// TIA Portal V21 export
// export: Created 2026-08-21T20:18:53.1493152Z, ExportSetting None, DisplayName Totally Integrated Automation Portal, DisplayVersion V21, DisplayName STEP 7 Professional, DisplayVersion V21, DisplayName STEP 7 Safety, DisplayVersion V21, DisplayName Tech WebApplication, DisplayVersion V21, DisplayName WinCC Basic/Comfort/Advanced, DisplayVersion V21, DisplayName WinCC Professional, DisplayVersion V21, DisplayName WinCC Unified, DisplayVersion V21
FUNCTION_BLOCK "ConfigurationParameters"   // FB1710, SCL
TITLE = ConfigurationParameters
{ S7_Optimized_Access := 'TRUE' }
AUTHOR : Siemens AG
FAMILY : ServiceControl
VERSION : 1.0
// Providing of the MTP-Interface and the number of parameters of each configuration parameter type
// stored: MemoryReserve 100, SetENOAutomatically false
   VAR
      MTPAnalog { S7_SetPoint := 'True'} : Array[0..#NUMBER_PARAMETERS_ANALOG] of "UDT_MTP_AnaServParam";
      MTPDigital { S7_SetPoint := 'True'} : Array[0..#NUMBER_PARAMETERS_DIGITAL] of "UDT_MTP_DIntServParam";
      MTPBinary { S7_SetPoint := 'True'} : Array[0..#NUMBER_PARAMETERS_BINARY] of "UDT_MTP_BinServParam";
      MTPString { S7_SetPoint := 'True'} : Array[0..#NUMBER_PARAMETERS_STRING] of "UDT_MTP_StringServParam";
   END_VAR
   VAR CONSTANT
      NUMBER_PARAMETERS_ANALOG : Int := 0;
      NUMBER_PARAMETERS_DIGITAL : Int := 0;
      NUMBER_PARAMETERS_BINARY : Int := 1;
      NUMBER_PARAMETERS_STRING : Int := 0;
   END_VAR
BEGIN
   REGION Block Info Header
     //===============================================================================
     // Siemens AG / (c)Copyright 2021
     //-------------------------------------------------------------------------------
     // Title:            ConfigurationParameters
     // Comment/Function: Providing of the MTP-Interface and the number of parameters of each configuration parameter type
     // Library/Family:   ServiceControl
     // Author:           Siemens AG
     // Tested with:      S7-PLCSIM Advanced 4.0
     // Engineering:      TIA Portal V17
     // Restrictions:     MTP
     // Requirements:     PLC (S7-1200 / S7-1500)
     //-------------------------------------------------------------------------------
     // Change log table:
     // Version  | Date       | Expert in charge        | Changes applied
     //----------|------------|-------------------------|-----------------------------
     // 01.00.00 | 02.09.2021 | Michael Schlosser       | First released version
     // 01.00.01 | 07.09.2021 | Michael Schlosser       | Change: Interface of FB28 ConfigurationParameterAnalog
     // 01.00.02 | 08.09.2021 | Michael Schlosser       | Change: Interface of FB18, FB33, FB24
     // 01.00.03 | 09.09.2021 | Michael Schlosser       | Change: For-loops only until #NUMBER_PARAMETERS_YXZ - 1
     // 01.00.04 | 15.09.2021 | Michael Schlosser       | Change: ApplyEn default values = true (e.g. parLevAnalogApplyEn[0])
     // 01.00.05 | 16.09.2021 | Michael Schlosser       | Change: ApplyEn & ApplyInt as part of UDT_Service_ParameterApply (e.g. #ParLevAnalogApply[0].En)
     // 01.00.06 | 18.10.2021 | Michael Schlosser       | change: call of FBs for parameters now in ServiceControlBlock-FBs to allow several services per PLC
     //===============================================================================
   END_REGION Block Info Header

   REGION Description
     // ConfigurationParameters provides the MTP-Interface and the number of parameters of each configuration parameter type
   END_REGION Description
END_FUNCTION_BLOCK
